Fanuc KAREL source: KD00005.KL

PROGRAM KD00005
%NOLOCKGROUP
%NOBUSYLAMP
VAR
  I: INTEGER
  J: INTEGER
  B: BOOLEAN
  R: REAL
  S: STRING[80]
BEGIN
  I = 1
END KD00005
